PROGRAM MAIN
VAR
	test : BOOL;
END_VAR

// Klopt dit?

END_PROGRAM

(* stored: Version 1.1.0.1
   POU MAIN: Id {8f50dd07-e275-4d5b-ba3f-83314db0c6b3}, SpecialFunc None *)
